// TIA Portal V20 export
TYPE "WT3_Kondensator_Status_UDT"
   STRUCT
      iHandshake : Int;
      Alarm : Struct
         bE0000_KonfigAlarm : Bool;
         bE0001_Reserviert : Bool;
         bE0002_InvUngueltig : Bool;
         bE0003_Reserviert : Bool;
         bE0004_Reserviert : Bool;
         bE0005_Reserviert : Bool;
         bE0006_WasserüberdruckZuTief : Bool;
         bE0007_Reserviert : Bool;
         bE0008_Reserviert : Bool;
         bE0009_Reserviert : Bool;
         bE0010_KondensatorpumpeAlarmBetrieb : Bool;
         bE0011_KondensatorpumpeAlarmStillstand : Bool;
         bE0012_KonfigAlarmVDMinVerflüssigungstemp : Bool;
         bE0013_KonfigAlarmCOPVerdichter : Bool;
         bE0014_DurchflussstörungKondImBetrieb : Bool;
         bE0015_DurchflussstörungKondIBeimStart : Bool;
         bE0016_DurchflussstörungKondImStillstand : Bool;
         bE0017_AbsperrklappeEintrittNichtOffen : Bool;
         bE0018_AbsperrklappeEintrittNichtZu : Bool;
         bE0019_AbsperrklappeAustrittNichtOffen : Bool;
         bE0020_AbsperrklappeAustrittNichtZu : Bool;
         bE0021_NH3inSekundärkreis : Bool;
         "bE0022_T-EintrittMaxblockiertVerdichterstart" : Bool;
         bE0023_StörungRegelventilAbscheider1 : Bool;
         bE0024_StörungRegelventilAbscheider2 : Bool;
         bE0025_ExternFehler : Bool;
         b052_Reserve : Bool;
         b053_Reserve : Bool;
         b054_Reserve : Bool;
         b055_Reserve : Bool;
         b056_Reserve : Bool;
         b057_Reserve : Bool;
         by06_Reserve : Byte;
         by07_Reserve : Byte;
         by08_Reserve : Byte;
         by09_Reserve : Byte;
         by10_Reserve : Byte;
         by11_Reserve : Byte;
         by12_Reserve : Byte;
         by13_Reserve : Byte;
         by14_Reserve : Byte;
         by15_Reserve : Byte;
         by16_Reserve : Byte;
         by17_Reserve : Byte;
         by18_Reserve : Byte;
         by19_Reserve : Byte;
         by20_Reserve : Byte;
         by21_Reserve : Byte;
         by22_Reserve : Byte;
         by23_Reserve : Byte;
         by24_Reserve : Byte;
         by25_Reserve : Byte;
         by26_Reserve : Byte;
         bE0200_AlarmKabelbruch : Bool;
         b271_Reserve : Bool;
         b272_Reserve : Bool;
         b273_Reserve : Bool;
         b274_Reserve : Bool;
         b275_Reserve : Bool;
         b276_Reserve : Bool;
         b277_Reserve : Bool;
         by28_Reserve : Byte;
         by29_Reserve : Byte;
         by30_Reserve : Byte;
         by31_Reserve : Byte;
         by32_Reserve : Byte;
         by33_Reserve : Byte;
      END_STRUCT;
      Warnung : Struct
         bA1000_Reserviert : Bool;
         bA1001_SlaveAusg : Bool;
         bA1002_Reserviert : Bool;
         bA1003_HauptMasterAusg : Bool;
         bA1004_MehrereKondensatorMasterAktiv : Bool;
         bA1005_ObjektIDMehrfachVorhanden : Bool;
         bA1006_Reserviert : Bool;
         bA1007_WassereingangstemperaturZuTief : Bool;
         bA1008_WarnungNiveauEndschalter : Bool;
         bA1009_WarnungNiveau2Endschalter : Bool;
         bA1010_Reserviert : Bool;
         bA1011_Reserviert : Bool;
         bA1012_Reserviert : Bool;
         bA1013_Reserviert : Bool;
         bA1014_Reserviert : Bool;
         bA1015_Reserviert : Bool;
         bA1016_Reserviert : Bool;
         b361_Reserve : Bool;
         b362_Reserve : Bool;
         b363_Reserve : Bool;
         b364_Reserve : Bool;
         b365_Reserve : Bool;
         b366_Reserve : Bool;
         b367_Reserve : Bool;
         by37_Reserve : Byte;
         by38_Reserve : Byte;
         by39_Reserve : Byte;
         by40_Reserve : Byte;
         by41_Reserve : Byte;
         by42_Reserve : Byte;
         by43_Reserve : Byte;
         by44_Reserve : Byte;
         by45_Reserve : Byte;
         by46_Reserve : Byte;
         by47_Reserve : Byte;
         by48_Reserve : Byte;
         by49_Reserve : Byte;
         by50_Reserve : Byte;
         by51_Reserve : Byte;
         by52_Reserve : Byte;
         by53_Reserve : Byte;
         by54_Reserve : Byte;
         by55_Reserve : Byte;
         by56_Reserve : Byte;
         by57_Reserve : Byte;
         by58_Reserve : Byte;
         bA1200_WarnungKabelbruch : Bool;
         b591_Reserve : Bool;
         b592_Reserve : Bool;
         b593_Reserve : Bool;
         b594_Reserve : Bool;
         b595_Reserve : Bool;
         b596_Reserve : Bool;
         b597_Reserve : Bool;
         by60_Reserve : Byte;
         by61_Reserve : Byte;
         by62_Reserve : Byte;
         by63_Reserve : Byte;
         by64_Reserve : Byte;
         by65_Reserve : Byte;
      END_STRUCT;
      Zustand : Struct
         bAlarmzustandAktiv : Bool;
         bWarnzustandAktiv : Bool;
         bSystemMeldungAktiv : Bool;
         bSeviceMeldungAktiv : Bool;
         bStopManuell : Bool;
         bStopAuto : Bool;
         bStopExtern : Bool;
         bBetriebAuto : Bool;
         bBetriebManuell : Bool;
         bAnlaufAuto : Bool;
         bAnlaufManuell : Bool;
         bManuellStoppen : Bool;
         b674_Reserve : Bool;
         b675_Reserve : Bool;
         b676_Reserve : Bool;
         b677_Reserve : Bool;
         by68_Reserve : Byte;
         by69_Reserve : Byte;
         bInventarAufnahme : Bool;
         b701_Reserve : Bool;
         bStandbyMasterInit : Bool;
         bStandbyMasterPassiv : Bool;
         bStandbyMasterAktiv : Bool;
         bNotbetriebAktiv : Bool;
         bMasterGesperrt : Bool;
         bSollwertAnhebung : Bool;
         bKondEintrittWarm : Bool;
         bIstwertVentilfühler : Bool;
         bIstwertPDruck : Bool;
         bKondensatorpumpeManuell : Bool;
         bAbsperrklappenOeffnen : Bool;
         bAbsperrklappenSchliessen : Bool;
         b716_Reserve : Bool;
         b717_Reserve : Bool;
         by72_Reserve : Byte;
         by73_Reserve : Byte;
         by74_Reserve : Byte;
         by75_Reserve : Byte;
         by76_Reserve : Byte;
         by77_Reserve : Byte;
         by78_Reserve : Byte;
         by79_Reserve : Byte;
         by80_Reserve : Byte;
         by81_Reserve : Byte;
      END_STRUCT;
      "Allgemeine Meldungen" : Struct
         b4000_AllgemeineMeldung_1 : Bool;
         b4001_AllgemeineMeldung_2 : Bool;
         b4002_AllgemeineMeldung_3 : Bool;
         b4003_AllgemeineMeldung_4 : Bool;
         b4004_AllgemeineMeldung_5 : Bool;
         b4005_AllgemeineMeldung_6 : Bool;
         b4006_AllgemeineMeldung_7 : Bool;
         b4007_AllgemeineMeldung_8 : Bool;
         by83_Reserve : Byte;
         by84_Reserve : Byte;
         by85_Reserve : Byte;
      END_STRUCT;
      DigIn : Struct
         b860_Reserve : Bool;
         bSollwertB : Bool;
         b862_Reserve : Bool;
         bNiveauregFreigabe : Bool;
         bNiveaureg2Freigabe : Bool;
         bWasserüberdruck : Bool;
         bNiveauEndschalterOffen : Bool;
         bNiveauEndschalterGeschlossen : Bool;
         bNiveau2EnschalterOffen : Bool;
         bNiveau2EnschalterGeschlossen : Bool;
         bEndschalterAbsperrklappeEintrittOffen : Bool;
         bEndschalterAbsperrklappeEintrittZu : Bool;
         bEndschalterAbsperrklappeAustrittOffen : Bool;
         bEndschalterAbsperrklappeAustrittZu : Bool;
         bNH3AlarmSekundärkreis : Bool;
         b877_Reserve : Bool;
         by88_Reserve : Byte;
         by89_Reserve : Byte;
         by90_Reserve : Byte;
         by91_Reserve : Byte;
         by92_Reserve : Byte;
         by93_Reserve : Byte;
      END_STRUCT;
      DigOut : Struct
         b940_Reserve : Bool;
         b941_Reserve : Bool;
         bKondensatorpumpe : Bool;
         bNiveauregelung : Bool;
         bNiveauregelung2 : Bool;
         bNiveauregelungDO : Bool;
         bNiveauregelung2DO : Bool;
         bAbsperrklappeEintritt : Bool;
         bAbsperrklappeAustritt : Bool;
         b951_Reserve : Bool;
         b952_Reserve : Bool;
         b953_Reserve : Bool;
         b954_Reserve : Bool;
         b955_Reserve : Bool;
         b956_Reserve : Bool;
         b957_Reserve : Bool;
         by96_Reserve : Byte;
         by97_Reserve : Byte;
         by98_Reserve : Byte;
         by99_Reserve : Byte;
         by100_Reserve : Byte;
         by101_Reserve : Byte;
      END_STRUCT;
      ch1021_Reserve : Char;
      chKondReglerEinheit : Char;
      rKondReglerIstwert : Real;
      rKondReglerSollwert : Real;
      rKondReglerAusgang : Real;
      rKondReglerStufen : Int;
      rKondEintrittstemperatur : Real;
      rKondAustrittstemperatur : Real;
      rAussentemperatur : Real;
      liSollwertUmschaltungStatus : DInt;
      rKondPISollwert : Real;
      rKondPIReglerIstwert : Real;
      rStellwert2Kd : Real;
      rKondensatorpumpe : Real;
      rKondDreiwegventil : Real;
      rFeuchtkugeltemperatur : Real;
      rT_Ventilfühler : Real;
      rNiveau : Real;
      rNiveauregulierung : Real;
      rNiveau2 : Real;
      rNiveauregulierung2 : Real;
      rVolumenstrom : Real;
      rThermischeLeistung : Real;
      rCOPVerdichter : Real;
      rCOPAnlage : Real;
      rWasserüberdruck : Real;
      rAuxAnalog1 : Real;
      rAuxAnalog2 : Real;
      rAuxAnalog3 : Real;
      rAuxAnalog4 : Real;
      byReserve : Array[214..629] of Byte;
   END_STRUCT;
END_TYPE
